FUNCTION_BLOCK Heating
VAR_INPUT
	diEnabled : BOOL;
	iSecImp : BOOL;
END_VAR
VAR_OUTPUT
	doEnabled : BOOL;
END_VAR
VAR_IN_OUT
	HeatingPhase : TPhaseHeating;
	Heater : THeater;
END_VAR
VAR
	pidParameters : ST_CTRL_PID_PARAMS;
	secImpTrig : R_TRIG;
END_VAR

{region "Aut/Man"}
    // switching state of engine - automatic or manual control (default state is manual)
    IF HeatingPhase.Cmd.ManCtrl THEN
        HeatingPhase.State.ManCtrl := TRUE;
        HeatingPhase.State.AutCtrl := FALSE;
    ELSIF HeatingPhase.Cmd.AutCtrl THEN
        HeatingPhase.State.ManCtrl := FALSE;
        HeatingPhase.State.AutCtrl := TRUE;
    END_IF;

    IF (NOT HeatingPhase.State.ManCtrl) AND (NOT HeatingPhase.State.AutCtrl) THEN
        HeatingPhase.State.ManCtrl := TRUE;
        HeatingPhase.State.AutCtrl := FALSE;
    END_IF;

    HeatingPhase.Cmd.ManCtrl := FALSE;
    HeatingPhase.Cmd.AutCtrl := FALSE;
{endregion}

{region "ManCtrl"}
    // processing manual actions - if command is processed, it is sets to FALSE even if can't be processed
    // real states of phase are writed into states in phase structure
    IF HeatingPhase.State.ManCtrl THEN
        IF HeatingPhase.Cmd.StartMan THEN
            HeatingPhase.State.Done := FALSE;
            IF HeatingPhase.State.Idle THEN
                HeatingPhase.fTime         := 0;
                HeatingPhase.State.Idle    := FALSE;
                HeatingPhase.State.Paused  := FALSE;
                HeatingPhase.State.Running := TRUE;
            END_IF;
        END_IF;

        IF HeatingPhase.Cmd.PauseMan THEN
            HeatingPhase.State.Done := FALSE;
            IF HeatingPhase.State.Running THEN
                HeatingPhase.State.Running := FALSE;
                HeatingPhase.State.Idle    := FALSE;
                HeatingPhase.State.Paused  := TRUE;
            END_IF;
        END_IF;

        IF HeatingPhase.Cmd.ResumeMan THEN
            HeatingPhase.State.Done := FALSE;
            IF HeatingPhase.State.Paused THEN
                HeatingPhase.State.Paused  := FALSE;
                HeatingPhase.State.Idle    := FALSE;
                HeatingPhase.State.Running := TRUE;
            END_IF;
        END_IF;

        IF HeatingPhase.Cmd.StopMan THEN
            HeatingPhase.State.Done    := FALSE;
            HeatingPhase.State.Running := FALSE;
            HeatingPhase.State.Paused  := FALSE;
            HeatingPhase.State.Idle    := TRUE;
            HeatingPhase.fTime         := 0;
        END_IF;
    END_IF;

    HeatingPhase.Cmd.StartMan  := FALSE;
    HeatingPhase.Cmd.StopMan   := FALSE;
    HeatingPhase.Cmd.PauseMan  := FALSE;
    HeatingPhase.Cmd.ResumeMan := FALSE;
{endregion}

{region "AutCtrl"}
    // if request to run in automatic mode -> set auto request to heat to 1, if not request to heat 0
    // commands should be sets to false after their processing
    IF HeatingPhase.State.AutCtrl THEN
        IF HeatingPhase.Cmd.StartAut THEN
            HeatingPhase.State.Done := FALSE;
            IF HeatingPhase.State.Idle THEN
                HeatingPhase.fTime         := 0;
                HeatingPhase.State.Idle    := FALSE;
                HeatingPhase.State.Paused  := FALSE;
                HeatingPhase.State.Running := TRUE;
            END_IF;
        END_IF;

        IF HeatingPhase.Cmd.StopAut THEN
            HeatingPhase.State.Done    := FALSE;
            HeatingPhase.State.Running := FALSE;
            HeatingPhase.State.Paused  := FALSE;
            HeatingPhase.State.Idle    := TRUE;
            HeatingPhase.fTime         := 0;
        END_IF;
    END_IF;

    HeatingPhase.Cmd.StartAut := FALSE;
    HeatingPhase.Cmd.StopAut  := FALSE;
{endregion}

{region "Done"}
    //every phase should have finish condition - heating phase - if water temp is on requested value for 10 seconds with 1°C hysteresis
    //after that done state should be setted to 1
    secImpTrig(CLK := iSecImp);

    IF HeatingPhase.State.Running THEN
        IF (HeatingPhase.WaterTemp >= (HeatingPhase.ParamReqTemp - 1.0)) AND (HeatingPhase.WaterTemp <= (HeatingPhase.ParamReqTemp + 1.0)) THEN
            IF secImpTrig.Q THEN
                HeatingPhase.fTime := HeatingPhase.fTime + 1;
            END_IF;
        ELSE
            HeatingPhase.fTime := 0;
        END_IF;

        IF HeatingPhase.fTime >= 1 THEN				/// TADY MA BYT 10
            HeatingPhase.State.Running := FALSE;
            HeatingPhase.State.Paused  := FALSE;
            HeatingPhase.State.Idle    := TRUE;
            HeatingPhase.State.Done    := TRUE;
            HeatingPhase.fTime         := 0;
        END_IF;
    ELSE
        HeatingPhase.fTime := 0;
    END_IF;

    // command reset done resets done state and than resets command
    IF HeatingPhase.Cmd.ResetDone THEN
        HeatingPhase.State.Done    := FALSE;
        HeatingPhase.Cmd.ResetDone := FALSE;
    END_IF;
{endregion}

{region "States"}
    //Command valve in cases of states
    // Running - start heating  
    // Idle - stop heating
    // Pause - stop heating (alternative is hold actual temp)
    IF HeatingPhase.State.Running THEN
        Heater.ParamHeatingSetPointAutomat := HeatingPhase.ParamReqTemp;
        Heater.Cmd.Req2RunAutCtrl := TRUE;
    ELSE
        Heater.Cmd.Req2RunAutCtrl := FALSE;
    END_IF;
{endregion}

// delault state of phase - if not any state sets state to idle
IF NOT HeatingPhase.State.Idle AND NOT HeatingPhase.State.Paused AND NOT HeatingPhase.State.Running THEN
    HeatingPhase.State.Idle := 1;
END_IF;

// write binary states into int value for visualization
IF HeatingPhase.State.Idle THEN
    HeatingPhase.State.Stateint := Global.PhIdle;
ELSIF HeatingPhase.State.Running THEN
    HeatingPhase.State.Stateint := Global.PhRunning;
ELSE
    HeatingPhase.State.Stateint := Global.PhPause;
END_IF;

doEnabled := diEnabled;

END_FUNCTION_BLOCK

(* stored: Version 1.1.0.1, ProductVersion 3.1.4026.21
   POU Heating: Id {67bfd793-3f9c-4f6b-ac3b-8ac7d5e1f5d7}, SpecialFunc None *)
